FUNCTION_BLOCK TANK_STRAPPING (* Migrated from IEC 61131-3 ST *)
  (* Standard: 61499-2 *)
  (* Version 1.0, 2026-11-06, st2fb *)
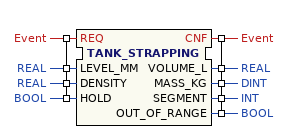
  EVENT_INPUT
    REQ WITH LEVEL_MM, DENSITY, HOLD;
  END_EVENT
  EVENT_OUTPUT
    CNF WITH VOLUME_L, MASS_KG, SEGMENT, OUT_OF_RANGE;
  END_EVENT
  VAR_INPUT
    LEVEL_MM : REAL;
    DENSITY : REAL;
    HOLD : BOOL;
  END_VAR
  VAR_OUTPUT
    VOLUME_L : REAL;
    MASS_KG : DINT;
    SEGMENT : INT;
    OUT_OF_RANGE : BOOL;
  END_VAR
  VAR
    L0 : REAL := 0.0;
    L1 : REAL := 200.0;
    L2 : REAL := 400.0;
    L3 : REAL := 800.0;
    L4 : REAL := 1200.0;
    L5 : REAL := 2000.0;
    V0 : REAL := 0.0;
    V1 : REAL := 150.0;
    V2 : REAL := 340.0;
    V3 : REAL := 800.0;
    V4 : REAL := 1350.0;
    V5 : REAL := 2600.0;
    I : INT := 0;
    FRACTION : REAL := 0.0;
    LA : REAL := 0.0;
    LB : REAL := 0.0;
    VA : REAL := 0.0;
    VB : REAL := 0.0;
    DONE : BOOL := FALSE;
  END_VAR
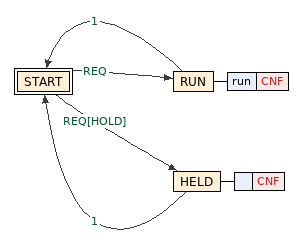
  EC_STATES
    START;
    RUN : run -> CNF;
    HELD : -> CNF;
  END_STATES
  EC_TRANSITIONS
    START TO HELD := REQ[HOLD];
    START TO RUN := REQ;
    RUN TO START := 1;
    HELD TO START := 1;
  END_TRANSITIONS
  ALGORITHM run IN ST:
OUT_OF_RANGE := (LEVEL_MM < L0) OR (LEVEL_MM > L5);
I := 0;
DONE := FALSE;
WHILE NOT DONE DO
  CASE I OF
    0: LB := L1;
    1: LB := L2;
    2: LB := L3;
    3: LB := L4;
    ELSE LB := L5;
  END_CASE;
  IF LEVEL_MM <= LB THEN
    DONE := TRUE;
  ELSE
    I := I + 1;
    IF I >= 4 THEN
      DONE := TRUE;
    END_IF;
  END_IF;
END_WHILE;
SEGMENT := I;
CASE I OF
  0: LA := L0; LB := L1; VA := V0; VB := V1;
  1: LA := L1; LB := L2; VA := V1; VB := V2;
  2: LA := L2; LB := L3; VA := V2; VB := V3;
  3: LA := L3; LB := L4; VA := V3; VB := V4;
  ELSE LA := L4; LB := L5; VA := V4; VB := V5;
END_CASE;
FRACTION := (LEVEL_MM - LA) / (LB - LA);
FRACTION := LIMIT(0.0, FRACTION, 1.0);
VOLUME_L := VA + FRACTION * (VB - VA);
MASS_KG := REAL_TO_DINT(VOLUME_L * DENSITY);
  END_ALGORITHM
END_FUNCTION_BLOCK
